Staubli VAL3: powerOnOff.pgx

public program powerOnOff(bool x_bPowerOn (dimensions=1))
begin
  if x_bPowerOn==true
    //Power on
    if !isPowered() and esStatus()!=2 and workingMode()==4
      autoConnectMove(true)
      enablePower()
      delay(1)
    endIf
  else
    //Power Off
    if isPowered()
      disablePower()
      delay(1)
    endIf
  endIf
end
